// I_Cabinet of the IAG50cm for the comm layer and the HMI gateway, with the physical Local/Remote key. The control mode is
// local while bLocalKey is TRUE and remote otherwise. Like FB_FixedCabinet, everything is an input of the block and there
// is no setter on I_Cabinet: the mode cannot become a software ownership switch over ADS, MQTT or the HMI.
FUNCTION_BLOCK FB_IagCabinet IMPLEMENTS I_Cabinet
VAR_INPUT
	bLocalKey			: BOOL;		// the Local/Remote key (FB_CabinetControl.LocalMode); TRUE = Local (polarity verified on site 2026-11-18: Remote reads 0, Local 1)
	bEstop				: BOOL;		// E-stop pressed or not yet released
	bSafetyError		: BOOL;		// TwinSAFE group in error
	bSafetyAckPending	: BOOL;		// E-stop released, acknowledge not run yet
	bPendantActive		: BOOL;		// a pendant holds motion authority
END_VAR

PROPERTY ControlMode : E_ControlMode
GET
ControlMode := SEL(bLocalKey, E_ControlMode.remote, E_ControlMode.local);
END_GET
END_PROPERTY

PROPERTY SwitchPresent : BOOL
GET
SwitchPresent := TRUE;
END_GET
END_PROPERTY

PROPERTY EstopActive : BOOL
GET
EstopActive := bEstop;
END_GET
END_PROPERTY

PROPERTY SafetyError : BOOL
GET
SafetyError := bSafetyError;
END_GET
END_PROPERTY

PROPERTY SafetyAckPending : BOOL
GET
SafetyAckPending := bSafetyAckPending;
END_GET
END_PROPERTY

PROPERTY PendantActive : BOOL
GET
PendantActive := bPendantActive;
END_GET
END_PROPERTY

END_FUNCTION_BLOCK

(* stored: Version 1.1.0.1, ProductVersion 3.1.4024.15
   POU FB_IagCabinet: Id {0af73759-ceed-421e-bb67-e4c267a398e7}, SpecialFunc None
   Property ControlMode: Id {989b5f90-4bc4-4926-8fd8-01e2823b7953}
   Get Get: Id {8e379851-e3bc-4cc3-905f-775300fb0343}
   Property SwitchPresent: Id {f618fcda-ea00-43a9-842a-0ecd1b26acde}
   Get Get: Id {a1dece7c-8509-4e1e-b4c5-e94fc1126cbd}
   Property EstopActive: Id {cf1ddcc9-d60f-4390-b8b3-24e54950c1b6}
   Get Get: Id {42f2cb1b-ab4f-4c26-a8c1-1586be79ce68}
   Property SafetyError: Id {14df7396-2676-4c14-9a7f-60216c8fac3d}
   Get Get: Id {09444a16-d9be-4a9f-8c96-258e701a461d}
   Property SafetyAckPending: Id {f58b446c-f55b-4fb2-8515-03e06d4dc75b}
   Get Get: Id {c471cda5-cf96-4e27-b999-6c3eda3059cd}
   Property PendantActive: Id {cc33a887-2004-43a2-b1ca-75555544a19f}
   Get Get: Id {ef27777f-2f4b-4055-a690-be2c85222a07} *)
